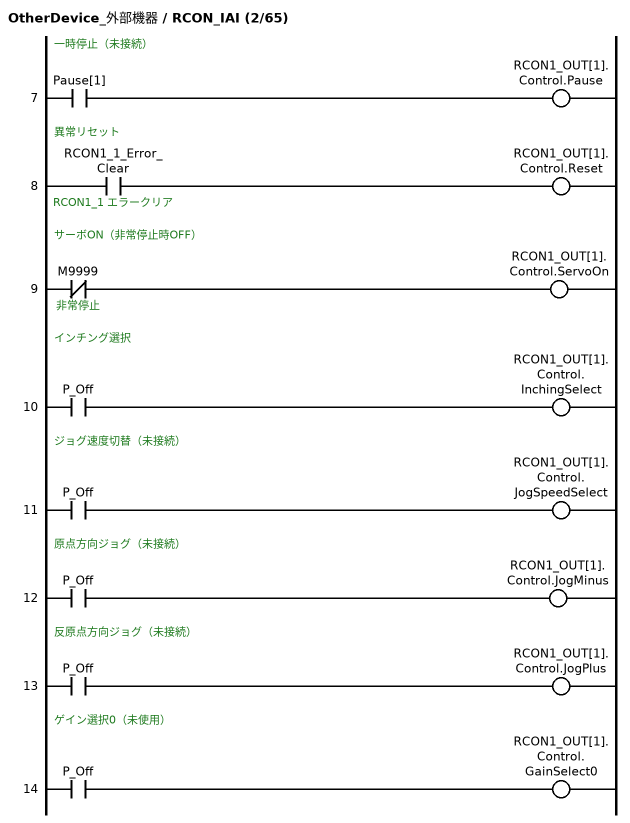
(* [picture p69: OtherDevice_外部機器 / RCON_IAI, rungs 7-14] *)
(* Rung 7: 一時停止（未接続） *)
RCON1_OUT[1].Control.Pause := Pause[1];
(* Rung 8: 異常リセット *)
RCON1_OUT[1].Control.Reset := RCON1_1_Error_Clear;
(* Rung 9: サーボON（非常停止時OFF） *)
RCON1_OUT[1].Control.ServoOn := NOT M9999;
(* Rung 10: インチング選択 *)
RCON1_OUT[1].Control.InchingSelect := P_Off;
(* Rung 11: ジョグ速度切替（未接続） *)
RCON1_OUT[1].Control.JogSpeedSelect := P_Off;
(* Rung 12: 原点方向ジョグ（未接続） *)
RCON1_OUT[1].Control.JogMinus := P_Off;
(* Rung 13: 反原点方向ジョグ（未接続） *)
RCON1_OUT[1].Control.JogPlus := P_Off;
(* Rung 14: ゲイン選択0（未使用） *)
RCON1_OUT[1].Control.GainSelect0 := P_Off;

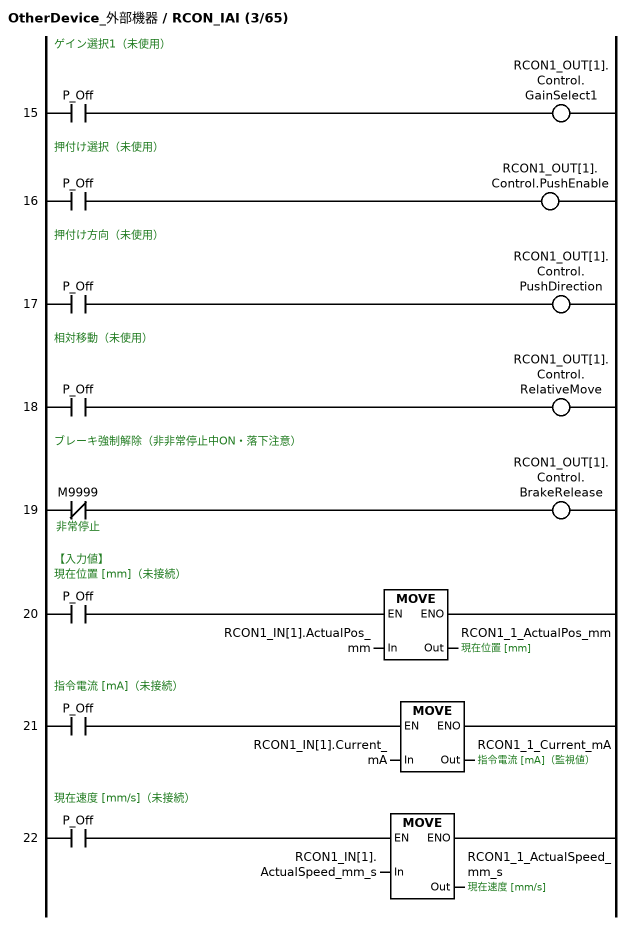
(* Rung 15: ゲイン選択1（未使用） *)
RCON1_OUT[1].Control.GainSelect1 := P_Off;
(* Rung 16: 押付け選択（未使用） *)
RCON1_OUT[1].Control.PushEnable := P_Off;
(* Rung 17: 押付け方向（未使用） *)
RCON1_OUT[1].Control.PushDirection := P_Off;
(* Rung 18: 相対移動（未使用） *)
RCON1_OUT[1].Control.RelativeMove := P_Off;
(* Rung 19: ブレーキ強制解除（非非常停止中ON・落下注意） *)
RCON1_OUT[1].Control.BrakeRelease := NOT M9999;
(* Rung 20: 【入力値】 / 現在位置 [mm]（未接続） *)
IF P_Off THEN RCON1_1_ActualPos_mm := RCON1_IN[1].ActualPos_mm; END_IF;
(* Rung 21: 指令電流 [mA]（未接続） *)
IF P_Off THEN RCON1_1_Current_mA := RCON1_IN[1].Current_mA; END_IF;
(* Rung 22: 現在速度 [mm/s]（未接続） *)
IF P_Off THEN RCON1_1_ActualSpeed_mm_s := RCON1_IN[1].ActualSpeed_mm_s; END_IF;

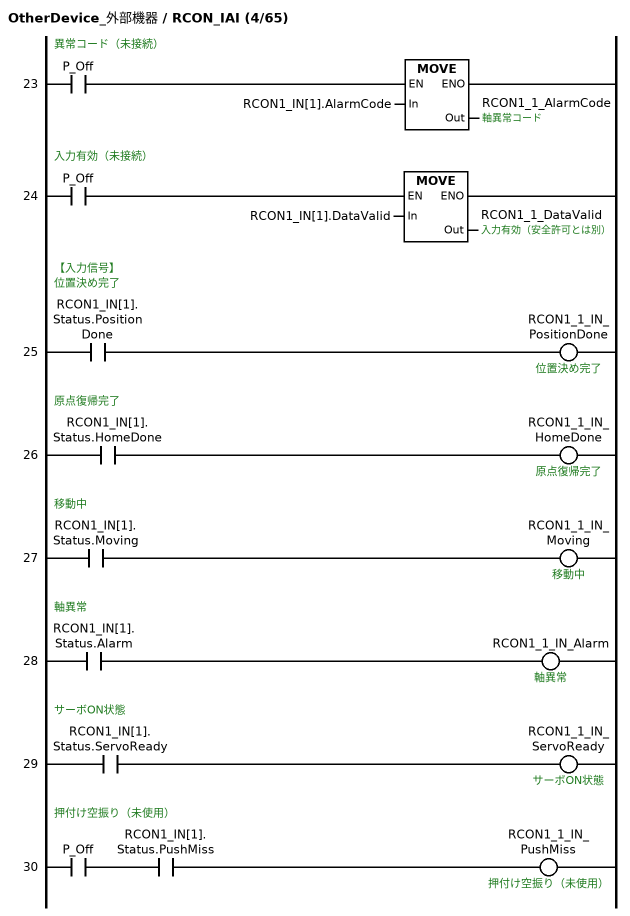
(* Rung 23: 異常コード（未接続） *)
IF P_Off THEN RCON1_1_AlarmCode := RCON1_IN[1].AlarmCode; END_IF;
(* Rung 24: 入力有効（未接続） *)
IF P_Off THEN RCON1_1_DataValid := RCON1_IN[1].DataValid; END_IF;
(* Rung 25: 【入力信号】 / 位置決め完了 *)
RCON1_1_IN_PositionDone := RCON1_IN[1].Status.PositionDone;
(* Rung 26: 原点復帰完了 *)
RCON1_1_IN_HomeDone := RCON1_IN[1].Status.HomeDone;
(* Rung 27: 移動中 *)
RCON1_1_IN_Moving := RCON1_IN[1].Status.Moving;
(* Rung 28: 軸異常 *)
RCON1_1_IN_Alarm := RCON1_IN[1].Status.Alarm;
(* Rung 29: サーボON状態 *)
RCON1_1_IN_ServoReady := RCON1_IN[1].Status.ServoReady;
(* Rung 30: 押付け空振り（未使用） *)
RCON1_1_IN_PushMiss := P_Off AND RCON1_IN[1].Status.PushMiss;

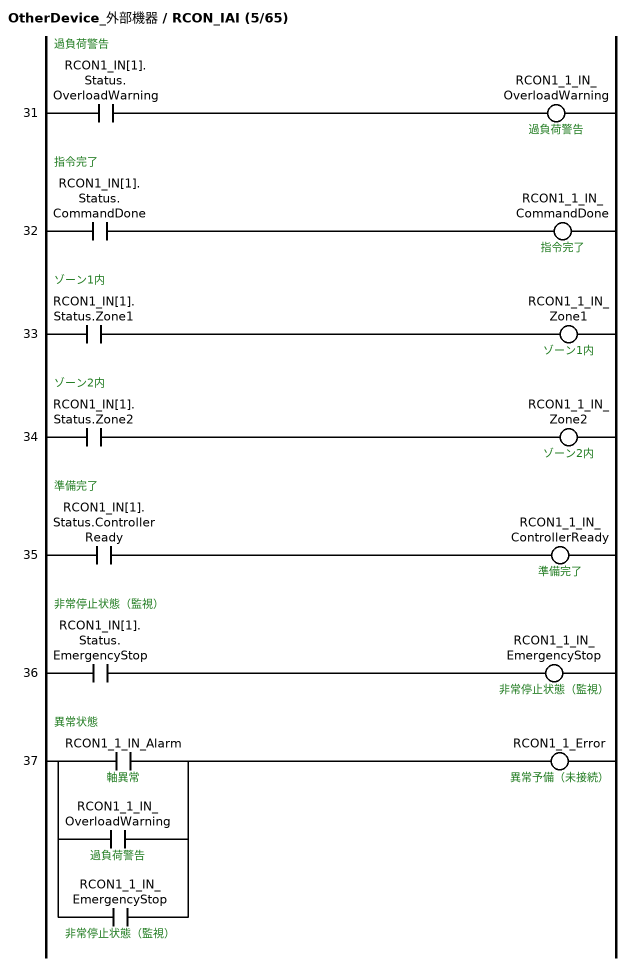
(* Rung 31: 過負荷警告 *)
RCON1_1_IN_OverloadWarning := RCON1_IN[1].Status.OverloadWarning;
(* Rung 32: 指令完了 *)
RCON1_1_IN_CommandDone := RCON1_IN[1].Status.CommandDone;
(* Rung 33: ゾーン1内 *)
RCON1_1_IN_Zone1 := RCON1_IN[1].Status.Zone1;
(* Rung 34: ゾーン2内 *)
RCON1_1_IN_Zone2 := RCON1_IN[1].Status.Zone2;
(* Rung 35: 準備完了 *)
RCON1_1_IN_ControllerReady := RCON1_IN[1].Status.ControllerReady;
(* Rung 36: 非常停止状態（監視） *)
RCON1_1_IN_EmergencyStop := RCON1_IN[1].Status.EmergencyStop;
(* Rung 37: 異常状態 *)
RCON1_1_Error := RCON1_1_IN_Alarm OR RCON1_1_IN_OverloadWarning OR RCON1_1_IN_EmergencyStop;

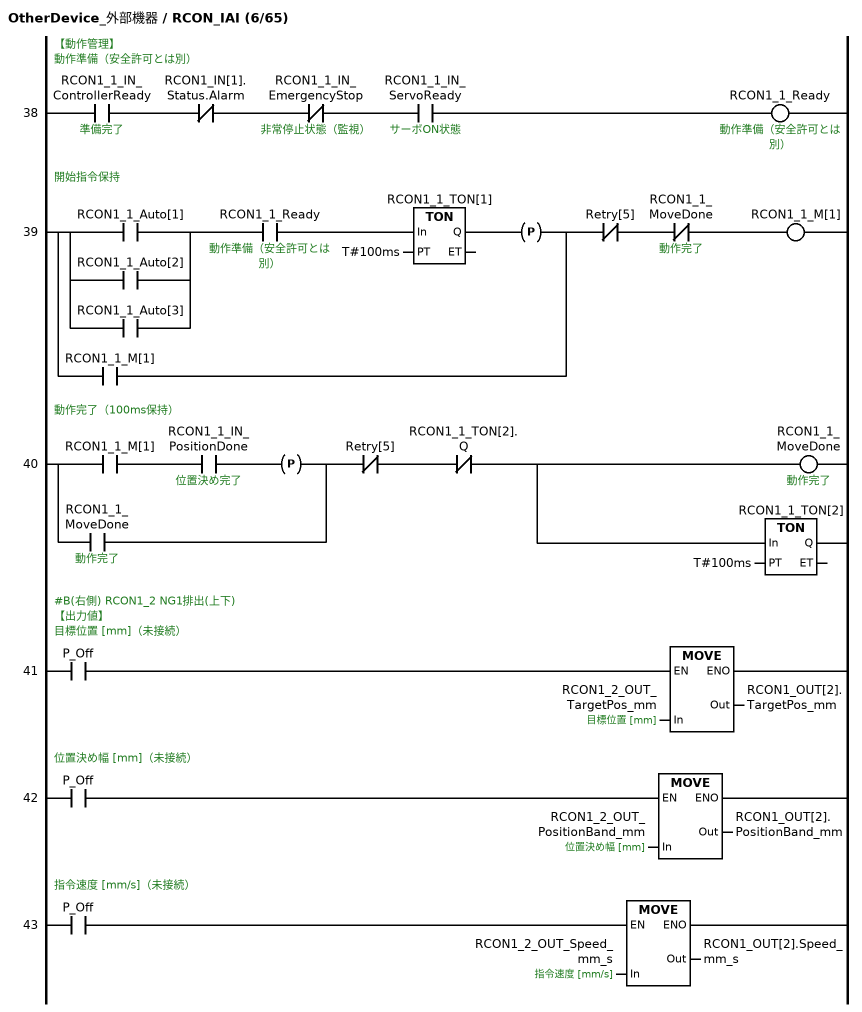
(* Rung 38: 【動作管理】 / 動作準備（安全許可とは別） *)
RCON1_1_Ready := RCON1_1_IN_ControllerReady AND NOT RCON1_IN[1].Status.Alarm AND NOT RCON1_1_IN_EmergencyStop AND RCON1_1_IN_ServoReady;
(* Rung 39: 開始指令保持 *)
RCON1_1_TON[1](In := (RCON1_1_Auto[1] OR RCON1_1_Auto[2] OR RCON1_1_Auto[3]) AND RCON1_1_Ready, PT := T#100ms);
_e2(CLK := RCON1_1_TON[1].Q);
RCON1_1_M[1] := (_e2.Q OR RCON1_1_M[1]) AND NOT Retry[5] AND NOT RCON1_1_MoveDone;
(* Rung 40: 動作完了（100ms保持） *)
_e3(CLK := RCON1_1_M[1] AND RCON1_1_IN_PositionDone);
_p4 := (_e3.Q OR RCON1_1_MoveDone) AND NOT Retry[5] AND NOT RCON1_1_TON[2].Q;
RCON1_1_MoveDone := _p4;
RCON1_1_TON[2](In := _p4, PT := T#100ms);
(* Rung 41: #B(右側) RCON1_2 NG1排出(上下) / 【出力値】 / 目標位置 [mm]（未接続） *)
IF P_Off THEN RCON1_OUT[2].TargetPos_mm := RCON1_2_OUT_TargetPos_mm; END_IF;
(* Rung 42: 位置決め幅 [mm]（未接続） *)
IF P_Off THEN RCON1_OUT[2].PositionBand_mm := RCON1_2_OUT_PositionBand_mm; END_IF;
(* Rung 43: 指令速度 [mm/s]（未接続） *)
IF P_Off THEN RCON1_OUT[2].Speed_mm_s := RCON1_2_OUT_Speed_mm_s; END_IF;

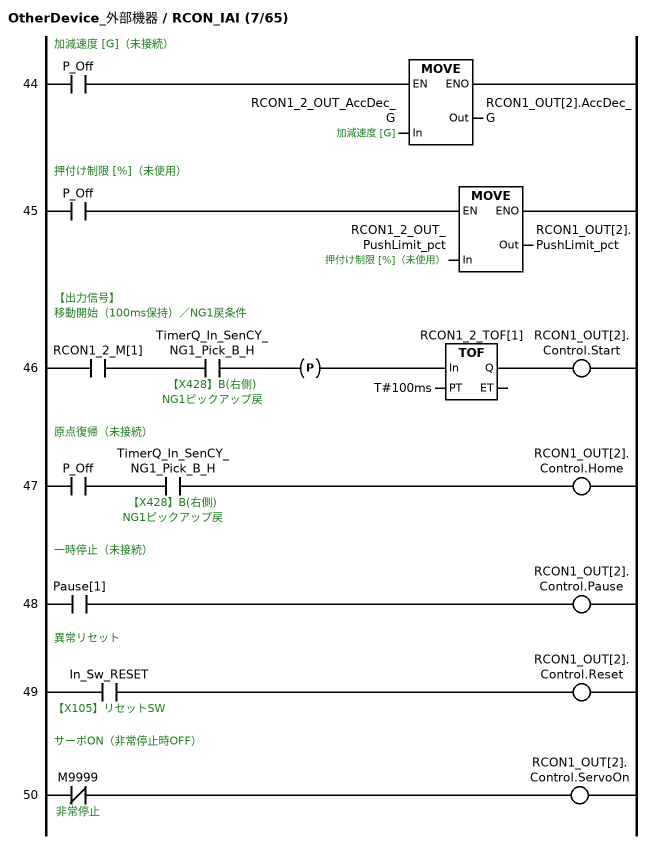
(* Rung 44: 加減速度 [G]（未接続） *)
IF P_Off THEN RCON1_OUT[2].AccDec_G := RCON1_2_OUT_AccDec_G; END_IF;
(* Rung 45: 押付け制限 [%]（未使用） *)
IF P_Off THEN RCON1_OUT[2].PushLimit_pct := RCON1_2_OUT_PushLimit_pct; END_IF;
(* Rung 46: 【出力信号】 / 移動開始（100ms保持）／NG1戻条件 *)
_e5(CLK := RCON1_2_M[1] AND TimerQ_In_SenCY_NG1_Pick_B_H);
RCON1_2_TOF[1](In := _e5.Q, PT := T#100ms);
RCON1_OUT[2].Control.Start := RCON1_2_TOF[1].Q;
(* Rung 47: 原点復帰（未接続） *)
RCON1_OUT[2].Control.Home := P_Off AND TimerQ_In_SenCY_NG1_Pick_B_H;
(* Rung 48: 一時停止（未接続） *)
RCON1_OUT[2].Control.Pause := Pause[1];
(* Rung 49: 異常リセット *)
RCON1_OUT[2].Control.Reset := In_Sw_RESET;
(* Rung 50: サーボON（非常停止時OFF） *)
RCON1_OUT[2].Control.ServoOn := NOT M9999;

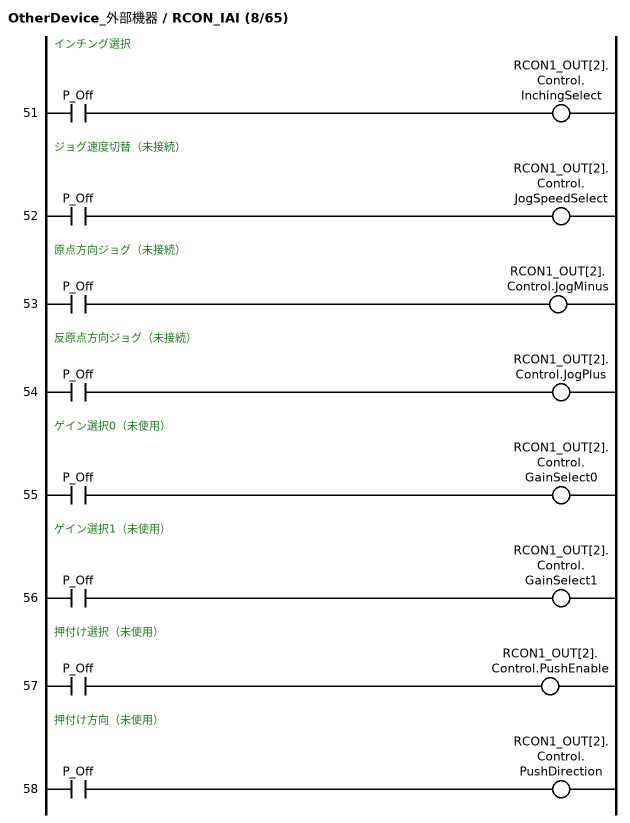
(* Rung 51: インチング選択 *)
RCON1_OUT[2].Control.InchingSelect := P_Off;
(* Rung 52: ジョグ速度切替（未接続） *)
RCON1_OUT[2].Control.JogSpeedSelect := P_Off;
(* Rung 53: 原点方向ジョグ（未接続） *)
RCON1_OUT[2].Control.JogMinus := P_Off;
(* Rung 54: 反原点方向ジョグ（未接続） *)
RCON1_OUT[2].Control.JogPlus := P_Off;
(* Rung 55: ゲイン選択0（未使用） *)
RCON1_OUT[2].Control.GainSelect0 := P_Off;
(* Rung 56: ゲイン選択1（未使用） *)
RCON1_OUT[2].Control.GainSelect1 := P_Off;
(* Rung 57: 押付け選択（未使用） *)
RCON1_OUT[2].Control.PushEnable := P_Off;
(* Rung 58: 押付け方向（未使用） *)
RCON1_OUT[2].Control.PushDirection := P_Off;

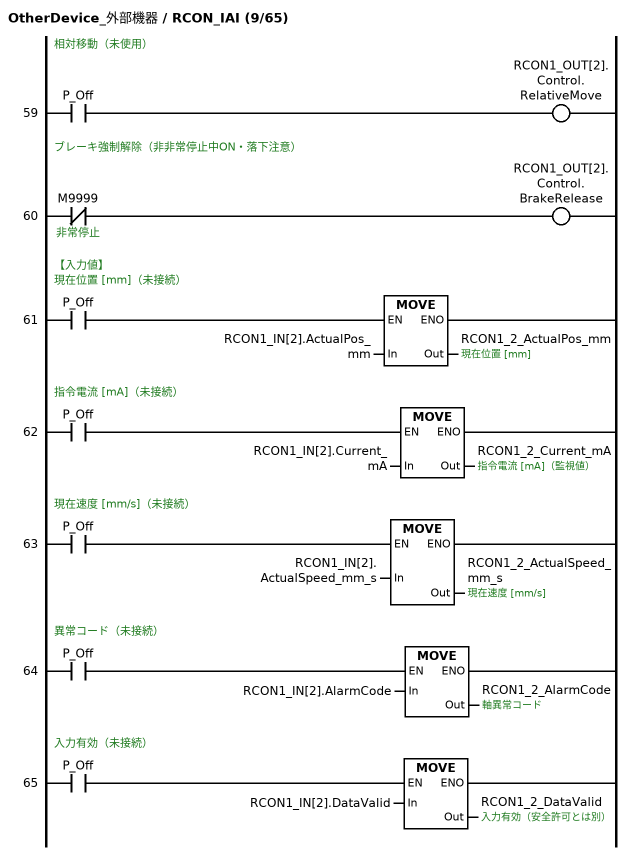
(* Rung 59: 相対移動（未使用） *)
RCON1_OUT[2].Control.RelativeMove := P_Off;
(* Rung 60: ブレーキ強制解除（非非常停止中ON・落下注意） *)
RCON1_OUT[2].Control.BrakeRelease := NOT M9999;
(* Rung 61: 【入力値】 / 現在位置 [mm]（未接続） *)
IF P_Off THEN RCON1_2_ActualPos_mm := RCON1_IN[2].ActualPos_mm; END_IF;
(* Rung 62: 指令電流 [mA]（未接続） *)
IF P_Off THEN RCON1_2_Current_mA := RCON1_IN[2].Current_mA; END_IF;
(* Rung 63: 現在速度 [mm/s]（未接続） *)
IF P_Off THEN RCON1_2_ActualSpeed_mm_s := RCON1_IN[2].ActualSpeed_mm_s; END_IF;
(* Rung 64: 異常コード（未接続） *)
IF P_Off THEN RCON1_2_AlarmCode := RCON1_IN[2].AlarmCode; END_IF;
(* Rung 65: 入力有効（未接続） *)
IF P_Off THEN RCON1_2_DataValid := RCON1_IN[2].DataValid; END_IF;

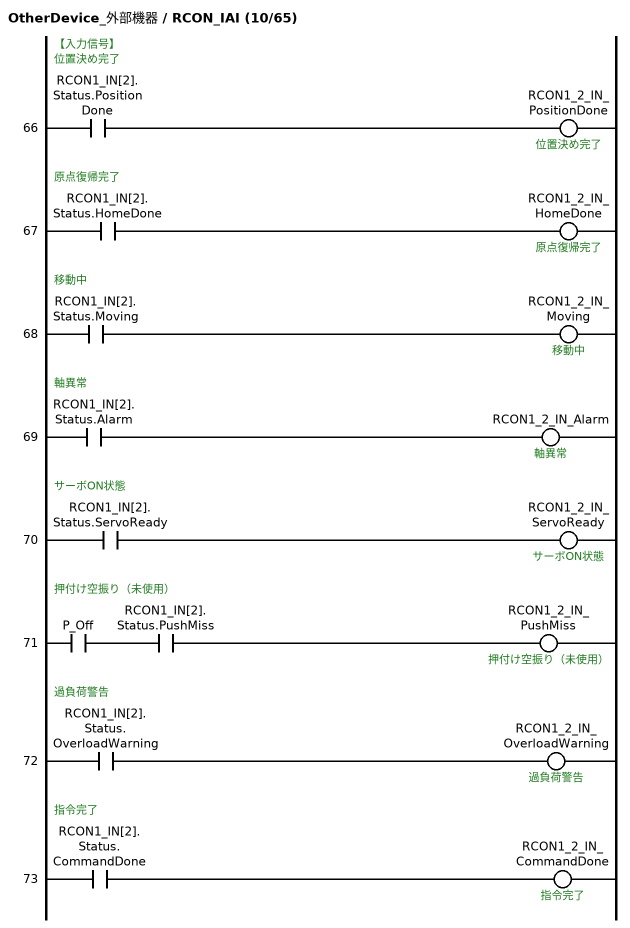
(* Rung 66: 【入力信号】 / 位置決め完了 *)
RCON1_2_IN_PositionDone := RCON1_IN[2].Status.PositionDone;
(* Rung 67: 原点復帰完了 *)
RCON1_2_IN_HomeDone := RCON1_IN[2].Status.HomeDone;
(* Rung 68: 移動中 *)
RCON1_2_IN_Moving := RCON1_IN[2].Status.Moving;
(* Rung 69: 軸異常 *)
RCON1_2_IN_Alarm := RCON1_IN[2].Status.Alarm;
(* Rung 70: サーボON状態 *)
RCON1_2_IN_ServoReady := RCON1_IN[2].Status.ServoReady;
(* Rung 71: 押付け空振り（未使用） *)
RCON1_2_IN_PushMiss := P_Off AND RCON1_IN[2].Status.PushMiss;
(* Rung 72: 過負荷警告 *)
RCON1_2_IN_OverloadWarning := RCON1_IN[2].Status.OverloadWarning;
(* Rung 73: 指令完了 *)
RCON1_2_IN_CommandDone := RCON1_IN[2].Status.CommandDone;

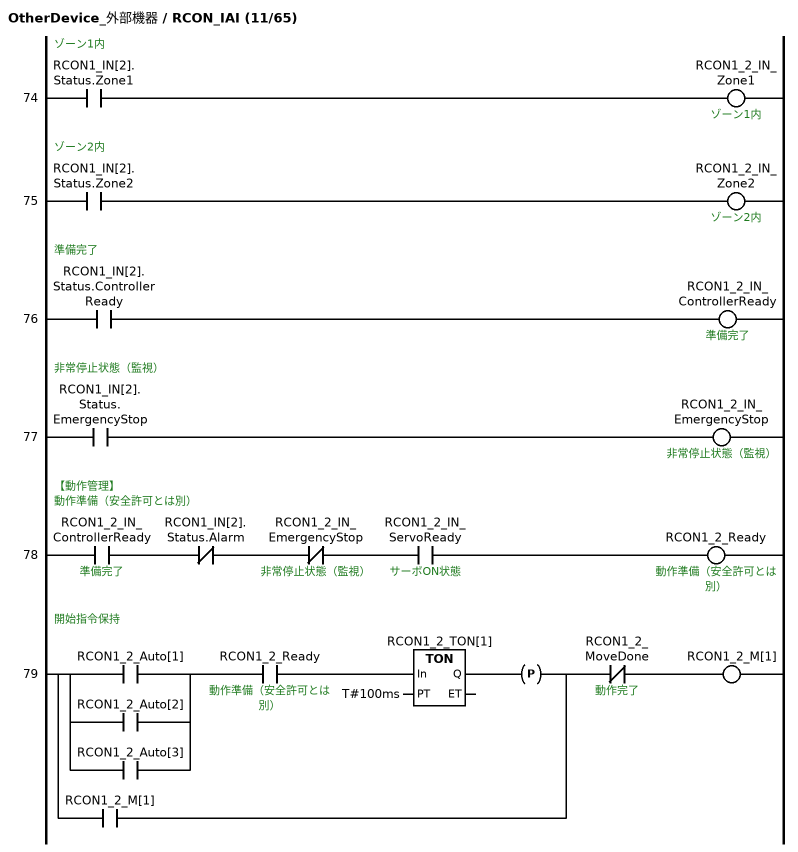
(* Rung 74: ゾーン1内 *)
RCON1_2_IN_Zone1 := RCON1_IN[2].Status.Zone1;
(* Rung 75: ゾーン2内 *)
RCON1_2_IN_Zone2 := RCON1_IN[2].Status.Zone2;
(* Rung 76: 準備完了 *)
RCON1_2_IN_ControllerReady := RCON1_IN[2].Status.ControllerReady;
(* Rung 77: 非常停止状態（監視） *)
RCON1_2_IN_EmergencyStop := RCON1_IN[2].Status.EmergencyStop;
(* Rung 78: 【動作管理】 / 動作準備（安全許可とは別） *)
RCON1_2_Ready := RCON1_2_IN_ControllerReady AND NOT RCON1_IN[2].Status.Alarm AND NOT RCON1_2_IN_EmergencyStop AND RCON1_2_IN_ServoReady;
(* Rung 79: 開始指令保持 *)
RCON1_2_TON[1](In := (RCON1_2_Auto[1] OR RCON1_2_Auto[2] OR RCON1_2_Auto[3]) AND RCON1_2_Ready, PT := T#100ms);
_e6(CLK := RCON1_2_TON[1].Q);
RCON1_2_M[1] := (_e6.Q OR RCON1_2_M[1]) AND NOT RCON1_2_MoveDone;

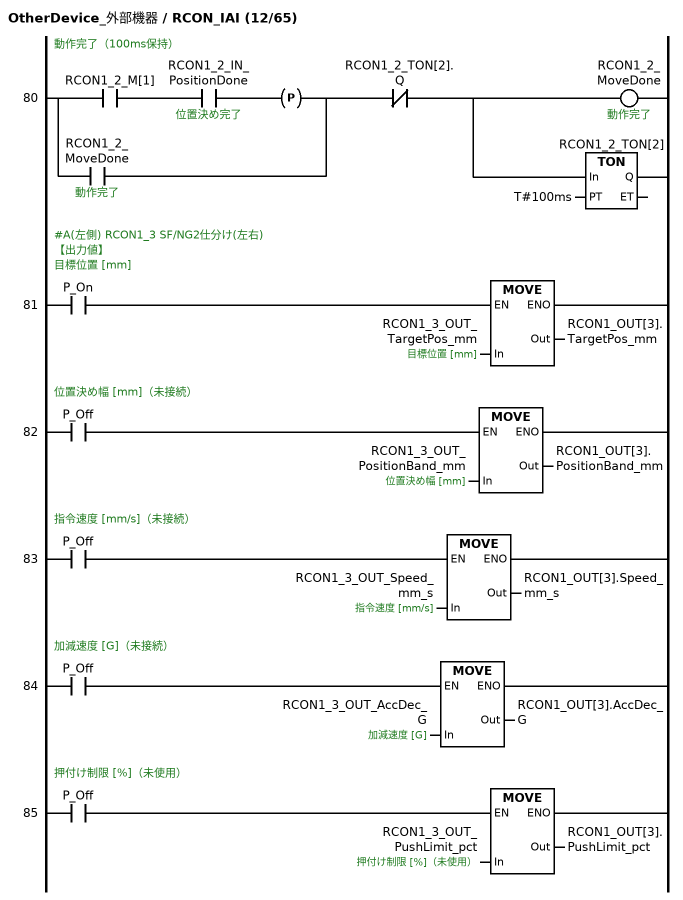
(* Rung 80: 動作完了（100ms保持） *)
_e7(CLK := RCON1_2_M[1] AND RCON1_2_IN_PositionDone);
_p8 := (_e7.Q OR RCON1_2_MoveDone) AND NOT RCON1_2_TON[2].Q;
RCON1_2_MoveDone := _p8;
RCON1_2_TON[2](In := _p8, PT := T#100ms);
(* Rung 81: #A(左側) RCON1_3 SF/NG2仕分け(左右) / 【出力値】 / 目標位置 [mm] *)
IF P_On THEN RCON1_OUT[3].TargetPos_mm := RCON1_3_OUT_TargetPos_mm; END_IF;
(* Rung 82: 位置決め幅 [mm]（未接続） *)
IF P_Off THEN RCON1_OUT[3].PositionBand_mm := RCON1_3_OUT_PositionBand_mm; END_IF;
(* Rung 83: 指令速度 [mm/s]（未接続） *)
IF P_Off THEN RCON1_OUT[3].Speed_mm_s := RCON1_3_OUT_Speed_mm_s; END_IF;
(* Rung 84: 加減速度 [G]（未接続） *)
IF P_Off THEN RCON1_OUT[3].AccDec_G := RCON1_3_OUT_AccDec_G; END_IF;
(* Rung 85: 押付け制限 [%]（未使用） *)
IF P_Off THEN RCON1_OUT[3].PushLimit_pct := RCON1_3_OUT_PushLimit_pct; END_IF;

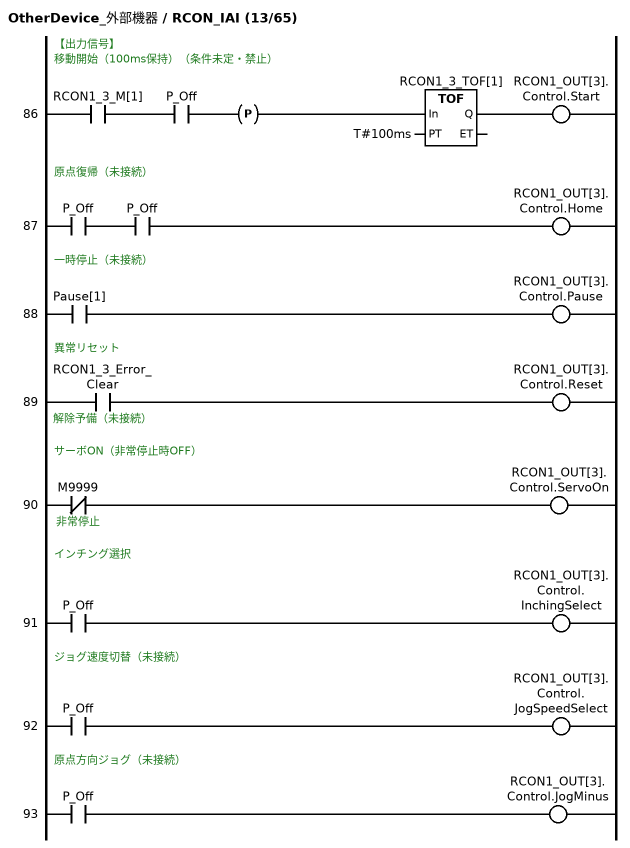
(* Rung 86: 【出力信号】 / 移動開始（100ms保持）（条件未定・禁止） *)
_e9(CLK := RCON1_3_M[1] AND P_Off);
RCON1_3_TOF[1](In := _e9.Q, PT := T#100ms);
RCON1_OUT[3].Control.Start := RCON1_3_TOF[1].Q;
(* Rung 87: 原点復帰（未接続） *)
RCON1_OUT[3].Control.Home := P_Off AND P_Off;
(* Rung 88: 一時停止（未接続） *)
RCON1_OUT[3].Control.Pause := Pause[1];
(* Rung 89: 異常リセット *)
RCON1_OUT[3].Control.Reset := RCON1_3_Error_Clear;
(* Rung 90: サーボON（非常停止時OFF） *)
RCON1_OUT[3].Control.ServoOn := NOT M9999;
(* Rung 91: インチング選択 *)
RCON1_OUT[3].Control.InchingSelect := P_Off;
(* Rung 92: ジョグ速度切替（未接続） *)
RCON1_OUT[3].Control.JogSpeedSelect := P_Off;
(* Rung 93: 原点方向ジョグ（未接続） *)
RCON1_OUT[3].Control.JogMinus := P_Off;

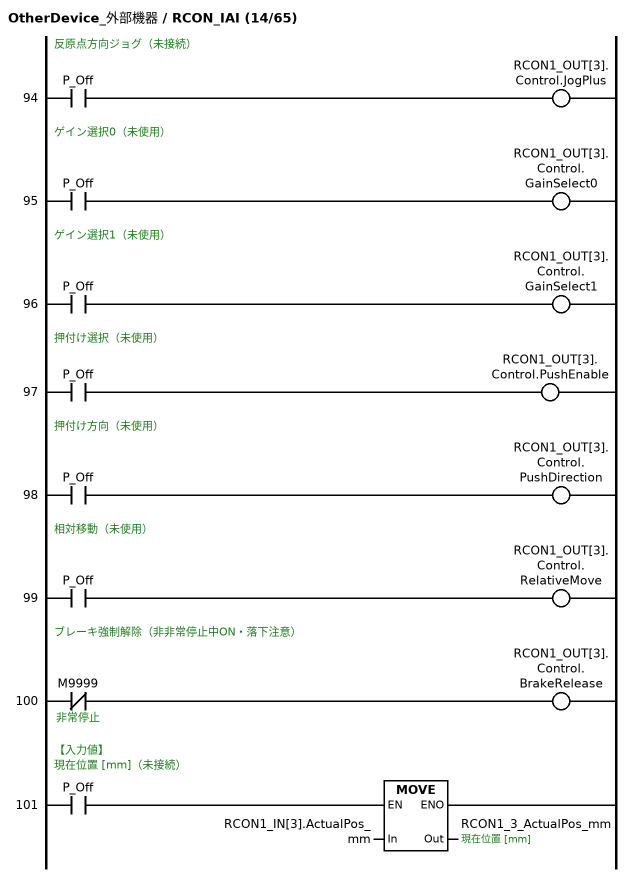
(* Rung 94: 反原点方向ジョグ（未接続） *)
RCON1_OUT[3].Control.JogPlus := P_Off;
(* Rung 95: ゲイン選択0（未使用） *)
RCON1_OUT[3].Control.GainSelect0 := P_Off;
(* Rung 96: ゲイン選択1（未使用） *)
RCON1_OUT[3].Control.GainSelect1 := P_Off;
(* Rung 97: 押付け選択（未使用） *)
RCON1_OUT[3].Control.PushEnable := P_Off;
(* Rung 98: 押付け方向（未使用） *)
RCON1_OUT[3].Control.PushDirection := P_Off;
(* Rung 99: 相対移動（未使用） *)
RCON1_OUT[3].Control.RelativeMove := P_Off;
(* Rung 100: ブレーキ強制解除（非非常停止中ON・落下注意） *)
RCON1_OUT[3].Control.BrakeRelease := NOT M9999;
(* Rung 101: 【入力値】 / 現在位置 [mm]（未接続） *)
IF P_Off THEN RCON1_3_ActualPos_mm := RCON1_IN[3].ActualPos_mm; END_IF;

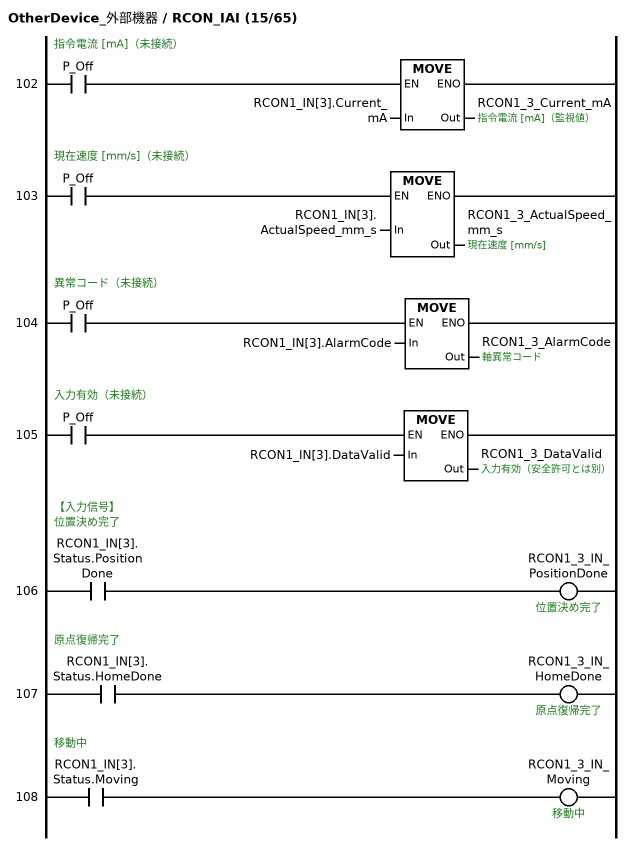
(* Rung 102: 指令電流 [mA]（未接続） *)
IF P_Off THEN RCON1_3_Current_mA := RCON1_IN[3].Current_mA; END_IF;
(* Rung 103: 現在速度 [mm/s]（未接続） *)
IF P_Off THEN RCON1_3_ActualSpeed_mm_s := RCON1_IN[3].ActualSpeed_mm_s; END_IF;
(* Rung 104: 異常コード（未接続） *)
IF P_Off THEN RCON1_3_AlarmCode := RCON1_IN[3].AlarmCode; END_IF;
(* Rung 105: 入力有効（未接続） *)
IF P_Off THEN RCON1_3_DataValid := RCON1_IN[3].DataValid; END_IF;
(* Rung 106: 【入力信号】 / 位置決め完了 *)
RCON1_3_IN_PositionDone := RCON1_IN[3].Status.PositionDone;
(* Rung 107: 原点復帰完了 *)
RCON1_3_IN_HomeDone := RCON1_IN[3].Status.HomeDone;
(* Rung 108: 移動中 *)
RCON1_3_IN_Moving := RCON1_IN[3].Status.Moving;

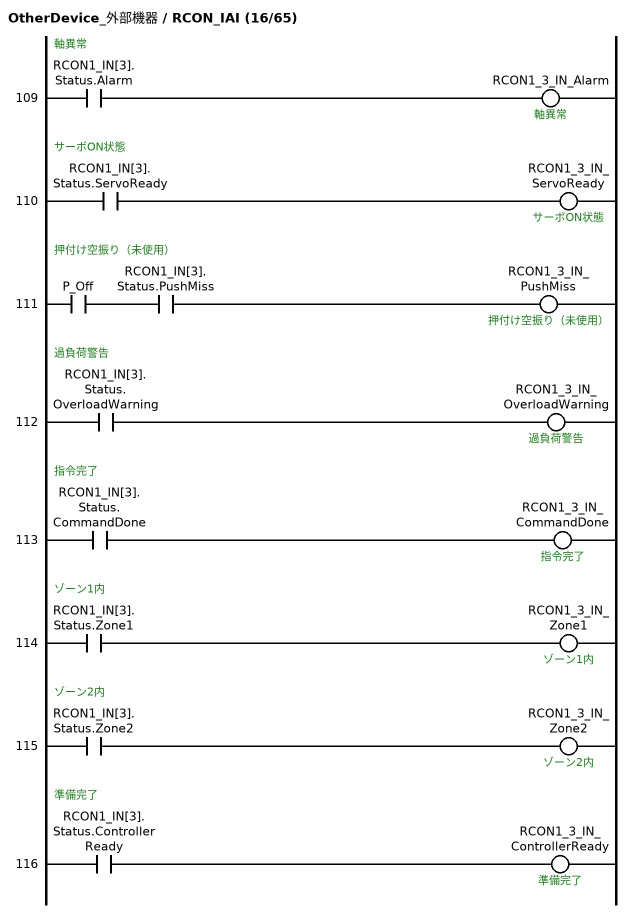
(* Rung 109: 軸異常 *)
RCON1_3_IN_Alarm := RCON1_IN[3].Status.Alarm;
(* Rung 110: サーボON状態 *)
RCON1_3_IN_ServoReady := RCON1_IN[3].Status.ServoReady;
(* Rung 111: 押付け空振り（未使用） *)
RCON1_3_IN_PushMiss := P_Off AND RCON1_IN[3].Status.PushMiss;
(* Rung 112: 過負荷警告 *)
RCON1_3_IN_OverloadWarning := RCON1_IN[3].Status.OverloadWarning;
(* Rung 113: 指令完了 *)
RCON1_3_IN_CommandDone := RCON1_IN[3].Status.CommandDone;
(* Rung 114: ゾーン1内 *)
RCON1_3_IN_Zone1 := RCON1_IN[3].Status.Zone1;
(* Rung 115: ゾーン2内 *)
RCON1_3_IN_Zone2 := RCON1_IN[3].Status.Zone2;
(* Rung 116: 準備完了 *)
RCON1_3_IN_ControllerReady := RCON1_IN[3].Status.ControllerReady;

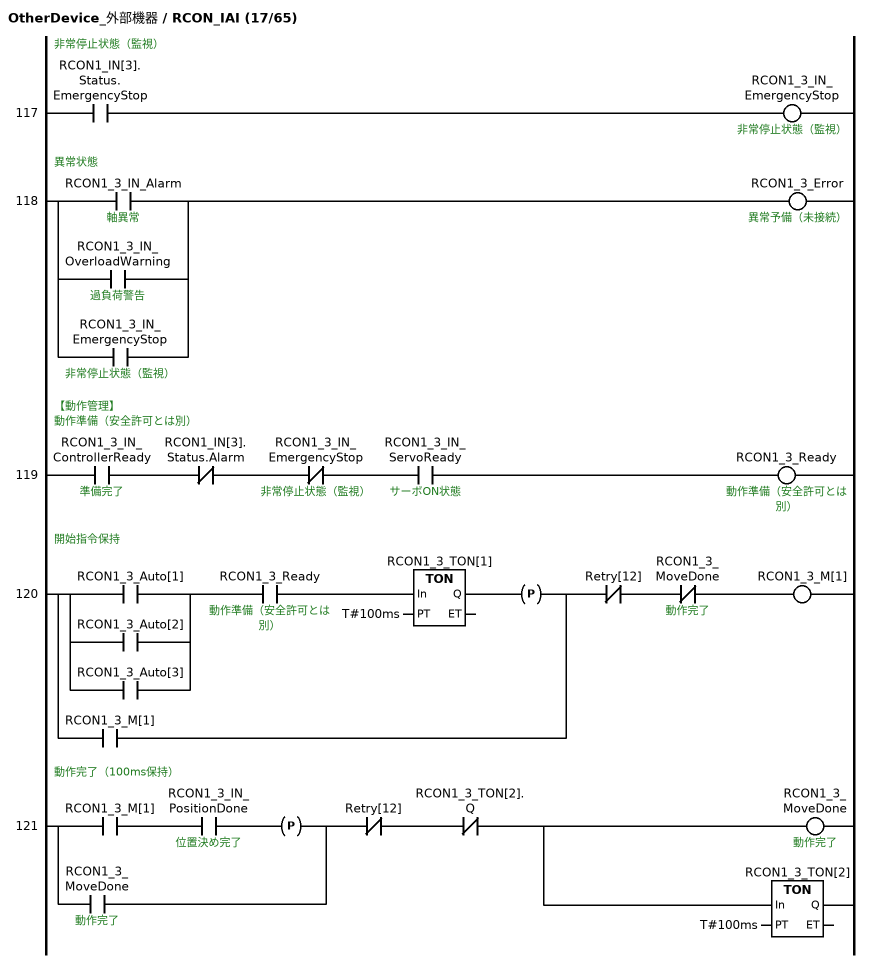
(* Rung 117: 非常停止状態（監視） *)
RCON1_3_IN_EmergencyStop := RCON1_IN[3].Status.EmergencyStop;
(* Rung 118: 異常状態 *)
RCON1_3_Error := RCON1_3_IN_Alarm OR RCON1_3_IN_OverloadWarning OR RCON1_3_IN_EmergencyStop;
(* Rung 119: 【動作管理】 / 動作準備（安全許可とは別） *)
RCON1_3_Ready := RCON1_3_IN_ControllerReady AND NOT RCON1_IN[3].Status.Alarm AND NOT RCON1_3_IN_EmergencyStop AND RCON1_3_IN_ServoReady;
(* Rung 120: 開始指令保持 *)
RCON1_3_TON[1](In := (RCON1_3_Auto[1] OR RCON1_3_Auto[2] OR RCON1_3_Auto[3]) AND RCON1_3_Ready, PT := T#100ms);
_e10(CLK := RCON1_3_TON[1].Q);
RCON1_3_M[1] := (_e10.Q OR RCON1_3_M[1]) AND NOT Retry[12] AND NOT RCON1_3_MoveDone;
(* Rung 121: 動作完了（100ms保持） *)
_e11(CLK := RCON1_3_M[1] AND RCON1_3_IN_PositionDone);
_p12 := (_e11.Q OR RCON1_3_MoveDone) AND NOT Retry[12] AND NOT RCON1_3_TON[2].Q;
RCON1_3_MoveDone := _p12;
RCON1_3_TON[2](In := _p12, PT := T#100ms);

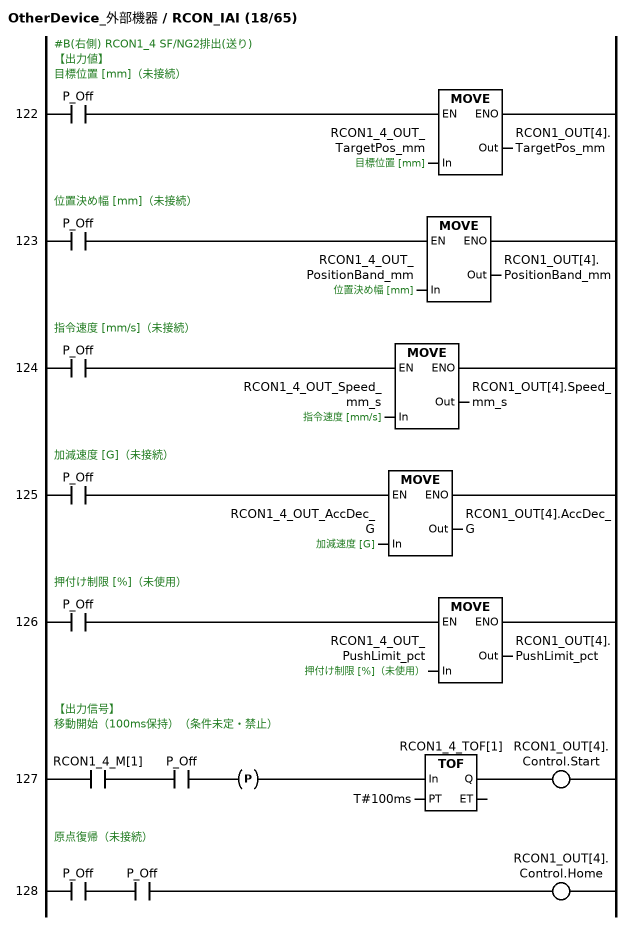
(* Rung 122: #B(右側) RCON1_4 SF/NG2排出(送り) / 【出力値】 / 目標位置 [mm]（未接続） *)
IF P_Off THEN RCON1_OUT[4].TargetPos_mm := RCON1_4_OUT_TargetPos_mm; END_IF;
(* Rung 123: 位置決め幅 [mm]（未接続） *)
IF P_Off THEN RCON1_OUT[4].PositionBand_mm := RCON1_4_OUT_PositionBand_mm; END_IF;
(* Rung 124: 指令速度 [mm/s]（未接続） *)
IF P_Off THEN RCON1_OUT[4].Speed_mm_s := RCON1_4_OUT_Speed_mm_s; END_IF;
(* Rung 125: 加減速度 [G]（未接続） *)
IF P_Off THEN RCON1_OUT[4].AccDec_G := RCON1_4_OUT_AccDec_G; END_IF;
(* Rung 126: 押付け制限 [%]（未使用） *)
IF P_Off THEN RCON1_OUT[4].PushLimit_pct := RCON1_4_OUT_PushLimit_pct; END_IF;
(* Rung 127: 【出力信号】 / 移動開始（100ms保持）（条件未定・禁止） *)
_e13(CLK := RCON1_4_M[1] AND P_Off);
RCON1_4_TOF[1](In := _e13.Q, PT := T#100ms);
RCON1_OUT[4].Control.Start := RCON1_4_TOF[1].Q;
(* Rung 128: 原点復帰（未接続） *)
RCON1_OUT[4].Control.Home := P_Off AND P_Off;

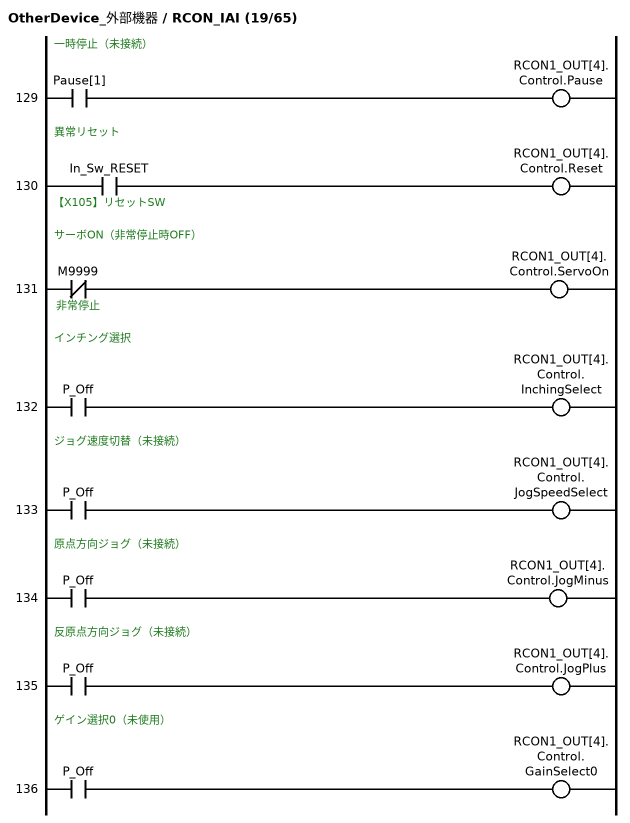
(* Rung 129: 一時停止（未接続） *)
RCON1_OUT[4].Control.Pause := Pause[1];
(* Rung 130: 異常リセット *)
RCON1_OUT[4].Control.Reset := In_Sw_RESET;
(* Rung 131: サーボON（非常停止時OFF） *)
RCON1_OUT[4].Control.ServoOn := NOT M9999;
(* Rung 132: インチング選択 *)
RCON1_OUT[4].Control.InchingSelect := P_Off;
(* Rung 133: ジョグ速度切替（未接続） *)
RCON1_OUT[4].Control.JogSpeedSelect := P_Off;
(* Rung 134: 原点方向ジョグ（未接続） *)
RCON1_OUT[4].Control.JogMinus := P_Off;
(* Rung 135: 反原点方向ジョグ（未接続） *)
RCON1_OUT[4].Control.JogPlus := P_Off;
(* Rung 136: ゲイン選択0（未使用） *)
RCON1_OUT[4].Control.GainSelect0 := P_Off;

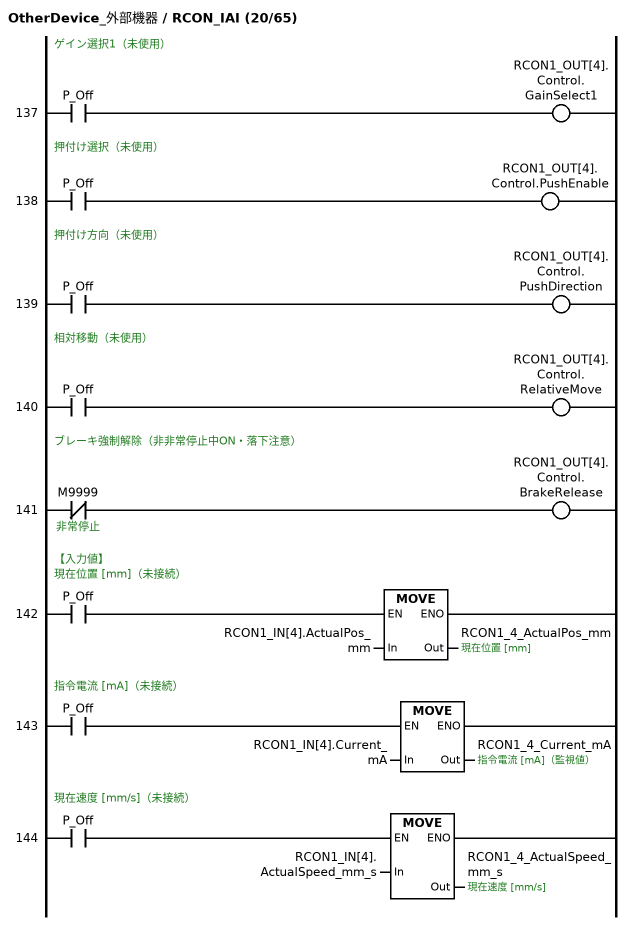
(* Rung 137: ゲイン選択1（未使用） *)
RCON1_OUT[4].Control.GainSelect1 := P_Off;
(* Rung 138: 押付け選択（未使用） *)
RCON1_OUT[4].Control.PushEnable := P_Off;
(* Rung 139: 押付け方向（未使用） *)
RCON1_OUT[4].Control.PushDirection := P_Off;
(* Rung 140: 相対移動（未使用） *)
RCON1_OUT[4].Control.RelativeMove := P_Off;
(* Rung 141: ブレーキ強制解除（非非常停止中ON・落下注意） *)
RCON1_OUT[4].Control.BrakeRelease := NOT M9999;
(* Rung 142: 【入力値】 / 現在位置 [mm]（未接続） *)
IF P_Off THEN RCON1_4_ActualPos_mm := RCON1_IN[4].ActualPos_mm; END_IF;
(* Rung 143: 指令電流 [mA]（未接続） *)
IF P_Off THEN RCON1_4_Current_mA := RCON1_IN[4].Current_mA; END_IF;
(* Rung 144: 現在速度 [mm/s]（未接続） *)
IF P_Off THEN RCON1_4_ActualSpeed_mm_s := RCON1_IN[4].ActualSpeed_mm_s; END_IF;

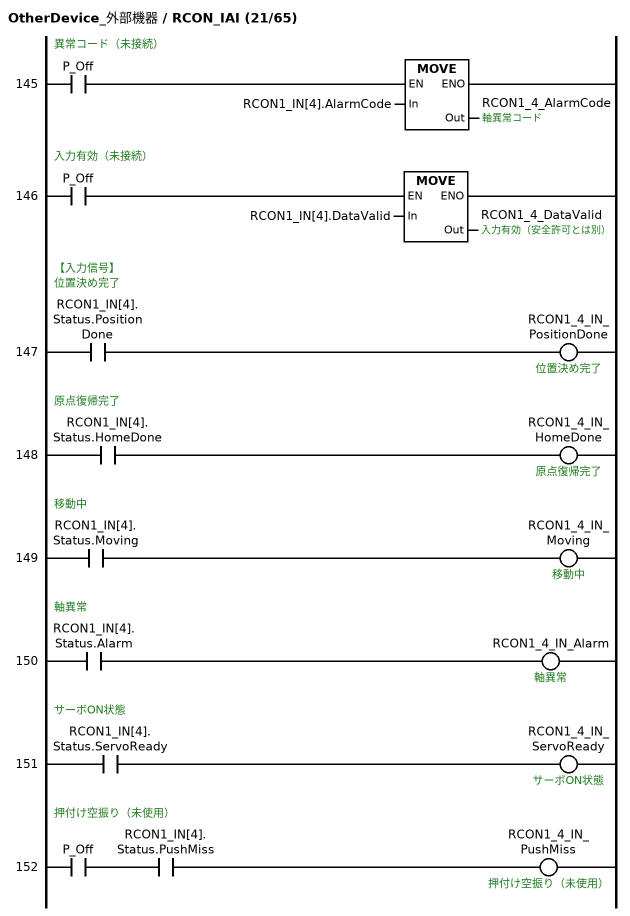
(* Rung 145: 異常コード（未接続） *)
IF P_Off THEN RCON1_4_AlarmCode := RCON1_IN[4].AlarmCode; END_IF;
(* Rung 146: 入力有効（未接続） *)
IF P_Off THEN RCON1_4_DataValid := RCON1_IN[4].DataValid; END_IF;
(* Rung 147: 【入力信号】 / 位置決め完了 *)
RCON1_4_IN_PositionDone := RCON1_IN[4].Status.PositionDone;
(* Rung 148: 原点復帰完了 *)
RCON1_4_IN_HomeDone := RCON1_IN[4].Status.HomeDone;
(* Rung 149: 移動中 *)
RCON1_4_IN_Moving := RCON1_IN[4].Status.Moving;
(* Rung 150: 軸異常 *)
RCON1_4_IN_Alarm := RCON1_IN[4].Status.Alarm;
(* Rung 151: サーボON状態 *)
RCON1_4_IN_ServoReady := RCON1_IN[4].Status.ServoReady;
(* Rung 152: 押付け空振り（未使用） *)
RCON1_4_IN_PushMiss := P_Off AND RCON1_IN[4].Status.PushMiss;

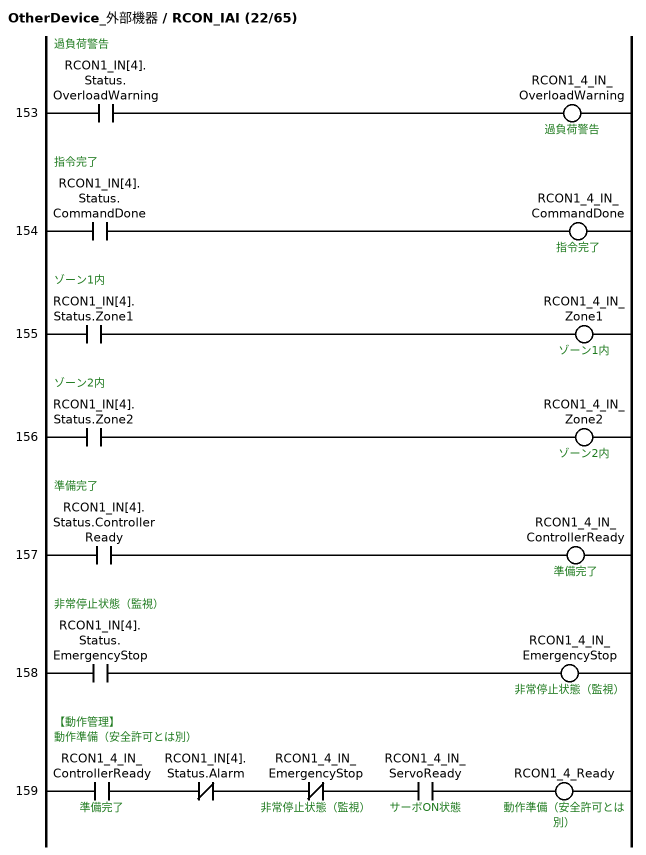
(* Rung 153: 過負荷警告 *)
RCON1_4_IN_OverloadWarning := RCON1_IN[4].Status.OverloadWarning;
(* Rung 154: 指令完了 *)
RCON1_4_IN_CommandDone := RCON1_IN[4].Status.CommandDone;
(* Rung 155: ゾーン1内 *)
RCON1_4_IN_Zone1 := RCON1_IN[4].Status.Zone1;
(* Rung 156: ゾーン2内 *)
RCON1_4_IN_Zone2 := RCON1_IN[4].Status.Zone2;
(* Rung 157: 準備完了 *)
RCON1_4_IN_ControllerReady := RCON1_IN[4].Status.ControllerReady;
(* Rung 158: 非常停止状態（監視） *)
RCON1_4_IN_EmergencyStop := RCON1_IN[4].Status.EmergencyStop;
(* Rung 159: 【動作管理】 / 動作準備（安全許可とは別） *)
RCON1_4_Ready := RCON1_4_IN_ControllerReady AND NOT RCON1_IN[4].Status.Alarm AND NOT RCON1_4_IN_EmergencyStop AND RCON1_4_IN_ServoReady;

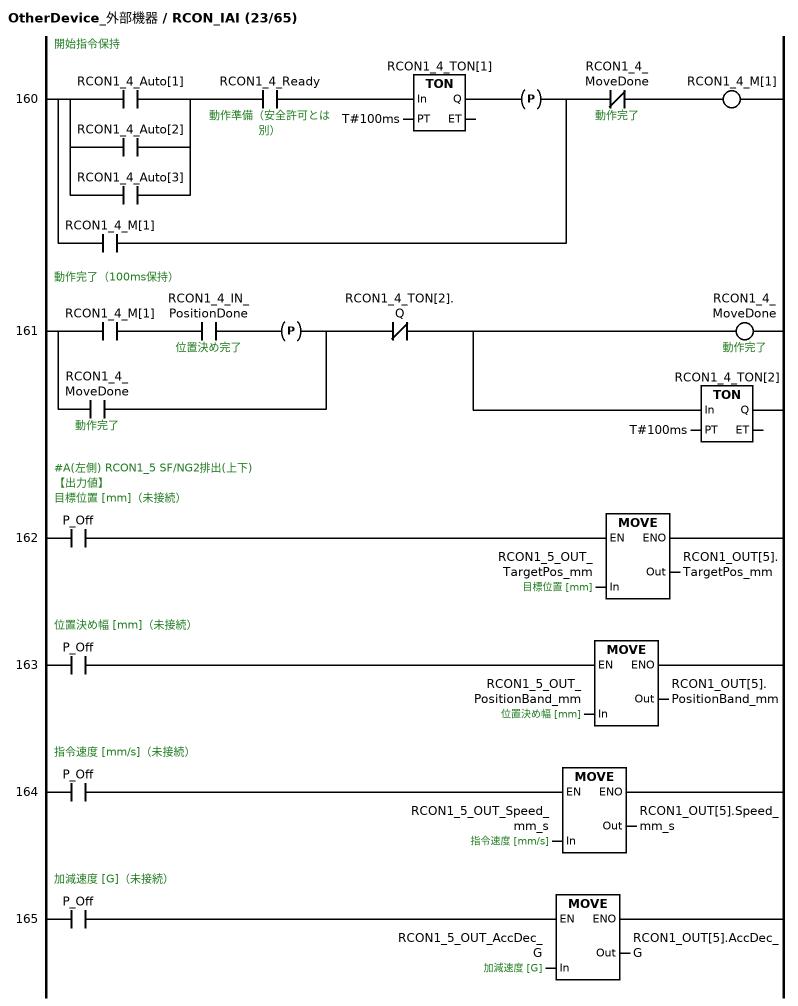
(* Rung 160: 開始指令保持 *)
RCON1_4_TON[1](In := (RCON1_4_Auto[1] OR RCON1_4_Auto[2] OR RCON1_4_Auto[3]) AND RCON1_4_Ready, PT := T#100ms);
_e14(CLK := RCON1_4_TON[1].Q);
RCON1_4_M[1] := (_e14.Q OR RCON1_4_M[1]) AND NOT RCON1_4_MoveDone;
(* Rung 161: 動作完了（100ms保持） *)
_e15(CLK := RCON1_4_M[1] AND RCON1_4_IN_PositionDone);
_p16 := (_e15.Q OR RCON1_4_MoveDone) AND NOT RCON1_4_TON[2].Q;
RCON1_4_MoveDone := _p16;
RCON1_4_TON[2](In := _p16, PT := T#100ms);
(* Rung 162: #A(左側) RCON1_5 SF/NG2排出(上下) / 【出力値】 / 目標位置 [mm]（未接続） *)
IF P_Off THEN RCON1_OUT[5].TargetPos_mm := RCON1_5_OUT_TargetPos_mm; END_IF;
(* Rung 163: 位置決め幅 [mm]（未接続） *)
IF P_Off THEN RCON1_OUT[5].PositionBand_mm := RCON1_5_OUT_PositionBand_mm; END_IF;
(* Rung 164: 指令速度 [mm/s]（未接続） *)
IF P_Off THEN RCON1_OUT[5].Speed_mm_s := RCON1_5_OUT_Speed_mm_s; END_IF;
(* Rung 165: 加減速度 [G]（未接続） *)
IF P_Off THEN RCON1_OUT[5].AccDec_G := RCON1_5_OUT_AccDec_G; END_IF;

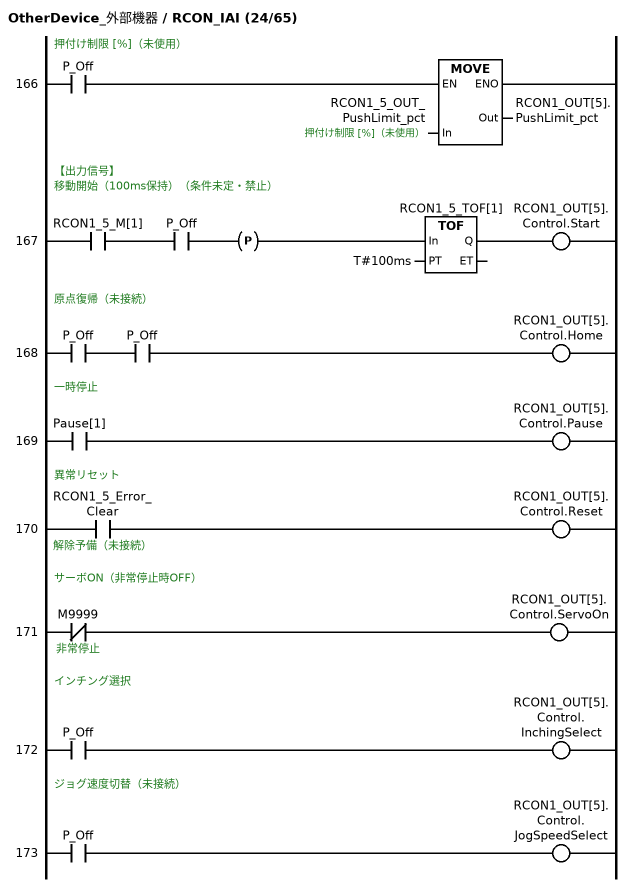
(* Rung 166: 押付け制限 [%]（未使用） *)
IF P_Off THEN RCON1_OUT[5].PushLimit_pct := RCON1_5_OUT_PushLimit_pct; END_IF;
(* Rung 167: 【出力信号】 / 移動開始（100ms保持）（条件未定・禁止） *)
_e17(CLK := RCON1_5_M[1] AND P_Off);
RCON1_5_TOF[1](In := _e17.Q, PT := T#100ms);
RCON1_OUT[5].Control.Start := RCON1_5_TOF[1].Q;
(* Rung 168: 原点復帰（未接続） *)
RCON1_OUT[5].Control.Home := P_Off AND P_Off;
(* Rung 169: 一時停止 *)
RCON1_OUT[5].Control.Pause := Pause[1];
(* Rung 170: 異常リセット *)
RCON1_OUT[5].Control.Reset := RCON1_5_Error_Clear;
(* Rung 171: サーボON（非常停止時OFF） *)
RCON1_OUT[5].Control.ServoOn := NOT M9999;
(* Rung 172: インチング選択 *)
RCON1_OUT[5].Control.InchingSelect := P_Off;
(* Rung 173: ジョグ速度切替（未接続） *)
RCON1_OUT[5].Control.JogSpeedSelect := P_Off;

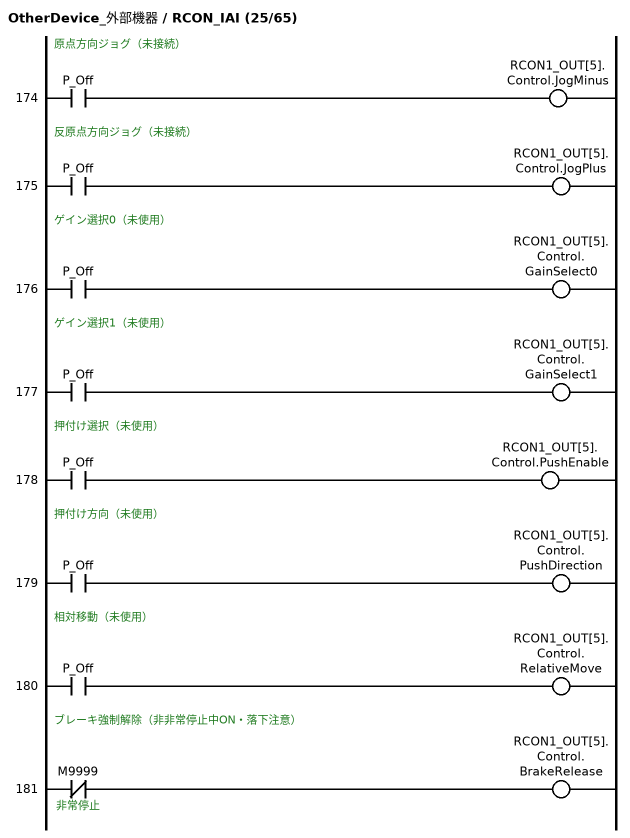
(* Rung 174: 原点方向ジョグ（未接続） *)
RCON1_OUT[5].Control.JogMinus := P_Off;
(* Rung 175: 反原点方向ジョグ（未接続） *)
RCON1_OUT[5].Control.JogPlus := P_Off;
(* Rung 176: ゲイン選択0（未使用） *)
RCON1_OUT[5].Control.GainSelect0 := P_Off;
(* Rung 177: ゲイン選択1（未使用） *)
RCON1_OUT[5].Control.GainSelect1 := P_Off;
(* Rung 178: 押付け選択（未使用） *)
RCON1_OUT[5].Control.PushEnable := P_Off;
(* Rung 179: 押付け方向（未使用） *)
RCON1_OUT[5].Control.PushDirection := P_Off;
(* Rung 180: 相対移動（未使用） *)
RCON1_OUT[5].Control.RelativeMove := P_Off;
(* Rung 181: ブレーキ強制解除（非非常停止中ON・落下注意） *)
RCON1_OUT[5].Control.BrakeRelease := NOT M9999;

